(*
SPDX-FileCopyrightText: c 2026 Oleksandr Tiutyk <trofimich@gmail.com>
SPDX-License-Identifier: MIT
License: https://opensource.org/license/mit
*)

(*!
<summary>Groups dynamic set lookup, duplicate updates, removal and clear cases.</summary>
<description>
Owns the child cases, their fixed registration array and the sets borrowed by the common cases.
Each borrowed fixture is reserved for its case throughout the group lifetime. Use from one task at a stable address.
</description>
*)

{attribute 'no_assign'}
{attribute 'no_explicit_call' := 'do not call this function block directly'}
FUNCTION_BLOCK DynamicUniqueDataSetTestGroup EXTENDS TOF_Testing.TestGroup<4>
VAR_STAT
	{attribute 'hide'}
	_ClassName : STRING := __POUNAME();
END_VAR
VAR
	_SetAndGetSet : TOF_Collections.UniqueDataSet<0>(valueValidator := 0, valueEqualityComparer := 0);
	_RemoveSet : TOF_Collections.UniqueDataSet<0>(valueValidator := 0, valueEqualityComparer := 0);
	_ContainsSet : TOF_Collections.UniqueDataSet<0>(valueValidator := 0, valueEqualityComparer := 0);

	_SetAndGet : UniqueDataSetSetAndGetTest(name := "SetAndGet", parent := THIS^, dataSet := _SetAndGetSet);
	_Remove : UniqueDataSetRemoveTest(name := "Remove", parent := THIS^, dataSet := _RemoveSet);
	_Contains : UniqueDataSetContainsTest(name := "Contains", parent := THIS^, dataSet := _ContainsSet);
	_Clear : DynamicUniqueDataSetClearTest(name := "Clear", parent := THIS^);

	_Children : ARRAY [0.._ChildCount - 1] OF TOF_Testing.ITestElement :=
	[
		_SetAndGet,
		_Remove,
		_Contains,
		_Clear
	];
END_VAR

//! <summary>Borrows the fixed child array. Callers must not modify it.</summary>
{attribute 'monitoring' := 'call'}
PROPERTY Children : REFERENCE TO ARRAY [0.._ChildCount - 1] OF TOF_Testing.ITestElement
GET
Children REF= _Children;
END_GET
END_PROPERTY

//! <summary>Borrows the concrete class name. Callers must not modify it.</summary>
{attribute 'monitoring' := 'call'}
PROPERTY ClassName : REFERENCE TO STRING
GET
ClassName REF= _ClassName;
END_GET
END_PROPERTY

//! <summary>Borrows the compiler-initialized namespace name. Callers must not modify it.</summary>
{attribute 'monitoring' := 'call'}
PROPERTY NamespaceName : REFERENCE TO STRING
GET
NamespaceName REF= CurrentNamespace.Name;
END_GET
END_PROPERTY

//! <summary>Reports the concrete instance size in bytes.</summary>
{attribute 'monitoring' := 'call'}
PROPERTY SelfSize : ULINT
GET
SelfSize := XSIZEOF(THIS^);
END_GET
END_PROPERTY

END_FUNCTION_BLOCK

(* stored: Version 1.1.0.1
   POU DynamicUniqueDataSetTestGroup: Id {6f389202-0508-41d6-adc8-91049d966d91}, SpecialFunc None
   Property Children: Id {80ee0d09-0f42-4631-b7ee-7d0106be9330}
   Get Get: Id {397a6b1d-1d8f-4c87-9e4a-844fd4b381fe}
   Property ClassName: Id {ce5fb722-4180-4d1f-a5f5-3cf0bb37fce6}
   Get Get: Id {bb0ef971-2c87-4ff6-baf0-6ac2e0a53b65}
   Property NamespaceName: Id {426e40ab-d79a-468f-b603-406767951b40}
   Get Get: Id {3e7b7908-e64b-4d7c-99bb-ef4dfd1d7bd4}
   Property SelfSize: Id {fa2d3f19-6312-47ad-b618-e018fd12dbf3}
   Get Get: Id {d3b22902-0402-43b3-a06f-86e0415bf3e7} *)
